FUNCTION_BLOCK T_SafeRs_Tests EXTENDS TcUnit.FB_TestSuite
VAR
    // Test_ResetDominantLatch
    group_1 : T_SafeGroup;
    fb_1 : T_SafeRs(group := group_1);
    // Test_UnconnectedSetIsRefused
    group_2 : T_SafeGroup;
    fb_2 : T_SafeRs(group := group_2);
END_VAR

Test_ResetDominantLatch();
Test_UnconnectedSetIsRefused();

METHOD PRIVATE Test_ResetDominantLatch
TcUnit.TEST(__POUNAME());
// act / assert
group_1(Run := TRUE);
fb_1(Set := TRUE, Reset := FALSE);
AssertEquals_BOOL(Expected := TRUE, Actual := fb_1.RsOut, Message := 'set');
fb_1(Set := FALSE, Reset := FALSE);
AssertEquals_BOOL(Expected := TRUE, Actual := fb_1.RsOut, Message := 'held');
fb_1(Set := TRUE, Reset := TRUE);
AssertEquals_BOOL(Expected := FALSE, Actual := fb_1.RsOut, Message := 'reset dominant');
TEST_FINISHED_NAMED(__POUNAME());
END_METHOD

METHOD PRIVATE Test_UnconnectedSetIsRefused
TcUnit.TEST(__POUNAME());
// arrange / act: Set is unconnected, which the Safety Editor refuses
group_2(Run := TRUE);
fb_2(Reset := FALSE);
group_2(Run := TRUE);
fb_2(Reset := FALSE);
// assert
AssertEquals_BOOL(Expected := TRUE, Actual := fb_2.Error, Message := 'configuration error reported');
AssertEquals_BYTE(Expected := TO_BYTE(E_SafeFbState.Error), Actual := fb_2.State, Message := 'state ERROR');
AssertEquals_WORD(Expected := WORD#16#8000, Actual := fb_2.Diag, Message := 'diag bit 15 configuration refused');
AssertEquals_BOOL(Expected := FALSE, Actual := fb_2.RsOut, Message := 'RsOut stays at its safe value');
AssertEquals_BOOL(Expected := TRUE, Actual := group_2.FbErr, Message := 'the group sees an FB error');
// act: ErrAck 0 -> 1 -> 0 does not clear a configuration error
group_2(Run := TRUE, ErrAck := TRUE);
fb_2(Reset := FALSE);
group_2(Run := TRUE, ErrAck := TRUE);
fb_2(Reset := FALSE);
group_2(Run := TRUE, ErrAck := FALSE);
fb_2(Reset := FALSE);
AssertEquals_BOOL(Expected := TRUE, Actual := fb_2.Error, Message := 'error not acknowledged');
AssertEquals_WORD(Expected := WORD#16#8000, Actual := fb_2.Diag, Message := 'diag bit 15 kept');
TEST_FINISHED_NAMED(__POUNAME());
END_METHOD

END_FUNCTION_BLOCK

(* stored: Version 1.1.0.1
   POU T_SafeRs_Tests: Id {292f3b71-3d46-58d8-a889-510872024b69}, SpecialFunc None
   Method Test_ResetDominantLatch: Id {d79316f9-bebc-55fe-a01d-0952a8c2e902}
   Method Test_UnconnectedSetIsRefused: Id {e2291759-74c8-4cd7-9edc-f2cc989bdf26} *)
